Fanuc KAREL source: NC0012.KL

PROGRAM NC0012
%NOLOCKGROUP
ROUTINE R
VAR
  X : INTEGER
BEGIN
  X = 1
  IF X = 1 THEN
    X = X + 2
  ELSE
    X = X + 1
  ENDIF
END R
BEGIN
  R
END NC0012
